TYPE E_VGC :
(

    Vented,
    AtVacuum,
    ERR_DiffPress,
    ERR_LostVac,
    ERR_ExtFault,
    At_Vac,
    Triggered,
    Vac_Fault,
    Cls_Timeout,
    Opn_Timeout


);
END_TYPE

(* stored: Version 1.1.0.1
   DUT E_VGC: Id {fcf967d4-478c-4b51-acfa-c0d70935d131} *)
